Fanuc KAREL source: kd00021.KL

-- PROVISIONAL review KL for V1013-1; original PC SHA256 39d02a54eca79254512dc4ce6f97e40f097260745b6ac09f47a401ca28da6787
-- Incomplete behavior may be omitted. Consult companion uncertainty JSON. Do not deploy.
PROGRAM KD00021
%NOLOCKGROUP
BEGIN
  -- UNRESOLVED_PC offsets 5-17; opcodes 21,23
  -- UNRESOLVED_PC offsets 22-26; opcodes 7F
END KD00021
